// TIA Portal project "交通灯 章家铭" (V15.1)

(* hardware
DEVICE "S7-1200 station_1"  S7-1200 Station
   slot 0: "Rack_0"  S7-1200 Rack  Rack  V1.0
   slot 1: "PLC_1"  CPU 1214C DC/DC/DC  6ES7 214-1AG40-0XB0  V4.2
   slot 2: "DI 16/DQ 16x24VDC_1"  6ES7 223-1BL32-0XB0  V2.0
   slot 3: "AI 4x13BIT/AQ 2x14BIT_1"  6ES7 234-4HE32-0XB0  V2.0
DEVICE "HMI_1"  KTP700 Basic PN
   slot 0: "HMI_1"  KTP700 Basic PN  6AV2 123-2GB03-0AX0  15.1.0.0
   slot 1: "HMI_RT_1"  KTP700 Basic PN  6AV2 123-2GB03-0AX0  15.1.0.0
   slot 5: "HMI_1.IE_CP_1"  PROFINET Interface  15.0.1.0
      slot 1: "PROFINET Interface_1"  PROFINET Interface
         slot 1: "Port_1"  Port
*)

// ===== PLC "PLC_1"  CPU 1214C DC/DC/DC =====

VAR_GLOBAL   // PLC tag table "默认变量表"
   "Tag_1" AT %I8.0 : Bool;
   "Tag_2" AT %I8.1 : Bool;
   "Tag_3" AT %I8.2 : Bool;
   "Tag_4" AT %I8.3 : Bool;
   "Tag_5" AT %I8.4 : Bool;
   "Tag_6" AT %I8.5 : Bool;
   "Tag_7" AT %I8.6 : Bool;
   "Tag_8" AT %I8.7 : Bool;
   "Tag_9" AT %I9.5 : Bool;
   "Tag_10" AT %Q8.0 : Bool;
   "Tag_11" AT %Q8.1 : Bool;
   "Tag_12" AT %Q8.2 : Bool;
   "Tag_13" AT %Q8.3 : Bool;
   "Tag_14" AT %Q8.4 : Bool;
   "Tag_15" AT %Q8.5 : Bool;
   "Tag_16" AT %Q8.6 : Bool;
   "Tag_17" AT %Q8.7 : Bool;
   "Tag_18" AT %Q9.0 : Bool;
   "Tag_19" AT %Q9.1 : Bool;
   "Tag_20" AT %Q9.2 : Bool;
   "Tag_21" AT %Q9.3 : Bool;
   "Tag_22" AT %Q9.4 : Bool;
   "Tag_23" AT %Q9.5 : Bool;
   "Tag_24" AT %Q9.6 : Bool;
   "Tag_25" AT %Q9.7 : Bool;
END_VAR

DATA_BLOCK "code_DB"   // DB1
{ S7_Optimized_Access := 'TRUE' }
VERSION : 0.1
// stored: InstanceOfName code
"code"
BEGIN
END_DATA_BLOCK

FUNCTION_BLOCK "code"   // FB1, SCL
{ S7_Optimized_Access := 'TRUE' }
VERSION : 0.1
   VAR_INPUT
      s01 : Bool;
      s02 : Bool;
      s03 : Bool;
      s04 : Bool;
      s05 : Bool;
      s06 : Bool;
      s07 : Bool;
      s14 : Bool;
   END_VAR
   VAR_OUTPUT
      k01 : Bool;
      k02 : Bool;
      k03 : Bool;
      k04 : Bool;
      k05 : Bool;
      k06 : Bool;
      k07 : Bool;
      k08 : Bool;
      k09 : Bool;
      k10 : Bool;
      k11 : Bool;
      k12 : Bool;
      k13 : Bool;
      k14 : Bool;
      k15 : Bool;
      k16 : Bool;
      hmi_ns_str_time : Int;
      hmi_ns_str_color : Int;
      hmi_ns_left_time : Int;
      hmi_ns_left_color : Int;
      hmi_ew_str_time : Int;
      hmi_ew_str_color : Int;
      hmi_ew_left_color : Int;
      hmi_ew_left_time : Int;
   END_VAR
   VAR
      auto_step : Int;
      ped_active : Bool;
      time_preset : Time;
      timer_auto : TON_TIME;
      timer_ped : TON_TIME;
   END_VAR
   VAR_TEMP
      elapsed_sec : Int;
      t_remain : Int;
      t_ped_remain : Int;
      blink_1hz : Bool;
   END_VAR
BEGIN
   // 初始化
   IF NOT #s01 THEN
       // 钥匙未开启时复位
       #auto_step := 0;
       #ped_active := FALSE;
   ELSE
       // 手动模式
       IF #s02 = TRUE THEN
           // 软件互锁：四个方向的绿灯请求互斥
           #k03 := #s03 AND NOT #s04 AND NOT #s05 AND NOT #s06;
           #k01 := NOT #k03;
           #k02 := FALSE;

           #k06 := #s04 AND NOT #s03 AND NOT #s05 AND NOT #s06;
           #k04 := NOT #k06;
           #k05 := FALSE;

           #k09 := #s05 AND NOT #s03 AND NOT #s04 AND NOT #s06;
           #k07 := NOT #k09;
           #k08 := FALSE;

           #k12 := #s06 AND NOT #s03 AND NOT #s04 AND NOT #s05;
           #k10 := NOT #k12;
           #k11 := FALSE;

           // 自动
       ELSE
           CASE #auto_step OF
               0:
                   #auto_step := 1;

               1:  // 南北直行绿灯
                   #time_preset := T#15s;
                   IF #timer_auto.Q THEN
                       #auto_step := 2;
                   END_IF;

               2:  // 南北直行黄灯
                   #time_preset := T#3s;
                   IF #timer_auto.Q THEN
                       #auto_step := 3;
                   END_IF;

               3:  // 南北左转绿灯
                   #time_preset := T#10s;
                   IF #timer_auto.Q THEN
                       #auto_step := 4;
                   END_IF;

               4:  // 南北左转黄灯
                   #time_preset := T#3s;
                   IF #timer_auto.Q THEN
                       #auto_step := 5;
                   END_IF;

               5:  // 东西直行绿灯
                   #time_preset := T#15s;
                   IF #timer_auto.Q THEN
                       #auto_step := 6;
                   END_IF;

               6:  // 东西直行黄灯
                   #time_preset := T#3s;
                   IF #timer_auto.Q THEN
                       #auto_step := 7;
                   END_IF;

               7:  // 东西左转绿灯
                   #time_preset := T#10s;
                   IF #timer_auto.Q THEN
                       #auto_step := 8;
                   END_IF;

               8:  // 东西左转黄灯
                   #time_preset := T#3s;
                   IF #timer_auto.Q THEN
                       #auto_step := 1;
                   END_IF;

               ELSE
                   #auto_step := 1;
           END_CASE;

           // 驱动自动模式的定时器
           #timer_auto(IN := TRUE,
                       PT := #time_preset);
           IF #timer_auto.Q THEN
               #timer_auto(IN := FALSE,
                           PT := #time_preset);
           END_IF;


           #blink_1hz := ((TIME_TO_DINT(#timer_auto.ET) / 500) MOD 2) = 0;

           #k03 := (#auto_step = 1);
           #k02 := (#auto_step = 2) AND #blink_1hz; 
           #k01 := NOT (#auto_step = 1 OR #auto_step = 2); 

           #k06 := (#auto_step = 3);
           #k05 := (#auto_step = 4) AND #blink_1hz;
           #k04 := NOT (#auto_step = 3 OR #auto_step = 4);

           #k09 := (#auto_step = 5);
           #k08 := (#auto_step = 6) AND #blink_1hz;
           #k07 := NOT (#auto_step = 5 OR #auto_step = 6);

           #k12 := (#auto_step = 7);
           #k11 := (#auto_step = 8) AND #blink_1hz;
           #k10 := NOT (#auto_step = 7 OR #auto_step = 8);


       END_IF;

       // 人行横道控制
       IF #s14 AND NOT #ped_active THEN
           #ped_active := TRUE;
       END_IF;

       // 行人过街定时逻辑
       #timer_ped(IN := #ped_active,
                  PT := T#5s);

       IF #ped_active THEN
           #k14 := FALSE;
           #k13 := TRUE;
           #k16 := FALSE;
           #k15 := TRUE;

           IF #timer_ped.Q THEN
               #ped_active := FALSE;
           END_IF;
       ELSE
           #k14 := TRUE;
           #k13 := FALSE;
           #k16 := TRUE;
           #k15 := FALSE;
       END_IF;

       // ==========================================
       // 5.倒计时
       // 颜色约定: 1=绿灯, 2=黄灯, 3=红灯
       // ==========================================
       IF #s02 THEN
           // 手动模式：没有倒计时(0)，只根据物理绿灯开关状态改变颜色
           #hmi_ns_str_time := 0;
           #hmi_ns_str_color := 3;
           IF #k03 THEN
               #hmi_ns_str_color := 1;
           END_IF;
           #hmi_ns_left_time := 0;
           #hmi_ns_left_color := 3;
           IF #k06 THEN
               #hmi_ns_left_color := 1;
           END_IF;
           #hmi_ew_str_time := 0;
           #hmi_ew_str_color := 3;
           IF #k09 THEN
               #hmi_ew_str_color := 1;
           END_IF;
           #hmi_ew_left_time := 0;
           #hmi_ew_left_color := 3;
           IF #k12 THEN
               #hmi_ew_left_color := 1;
           END_IF;
       ELSE
           // 自动模式：提取当前相位剩余的秒数
           #t_remain := DINT_TO_INT(TIME_TO_DINT(#time_preset) / 1000) - DINT_TO_INT(TIME_TO_DINT(#timer_auto.ET) / 1000);
           IF #t_remain < 0 THEN
               #t_remain := 0;
           END_IF;

           // 核心时间轴投射 (精确计算其他方向等待绿灯的时间)
           CASE #auto_step OF
               1: // 相位: 南北直行绿灯
                   #hmi_ns_str_time := #t_remain;
                   #hmi_ns_str_color := 1; // 绿
                   #hmi_ns_left_time := #t_remain + 3;
                   #hmi_ns_left_color := 3; // 红 (等接下来的黄灯走完)
                   #hmi_ew_str_time := #t_remain + 16;
                   #hmi_ew_str_color := 3; // 红 (3黄+10左+3黄)
                   #hmi_ew_left_time := #t_remain + 34;
                   #hmi_ew_left_color := 3; // 红
               2: // 相位: 南北直行黄灯
                   #hmi_ns_str_time := #t_remain;
                   #hmi_ns_str_color := 2; // 黑
                   #hmi_ns_left_time := #t_remain;
                   #hmi_ns_left_color := 3;
                   #hmi_ew_str_time := #t_remain + 13;
                   #hmi_ew_str_color := 3;
                   #hmi_ew_left_time := #t_remain + 31;
                   #hmi_ew_left_color := 3;
               3: // 相位: 南北左转绿灯
                   #hmi_ns_str_time := #t_remain + 34;
                   #hmi_ns_str_color := 3; // 红
                   #hmi_ns_left_time := #t_remain;
                   #hmi_ns_left_color := 1; // 绿
                   #hmi_ew_str_time := #t_remain + 3;
                   #hmi_ew_str_color := 3;
                   #hmi_ew_left_time := #t_remain + 21;
                   #hmi_ew_left_color := 3;
               4: // 相位: 南北左转黄灯
                   #hmi_ns_str_time := #t_remain + 31;
                   #hmi_ns_str_color := 3;
                   #hmi_ns_left_time := #t_remain;
                   #hmi_ns_left_color := 2; // 黑
                   #hmi_ew_str_time := #t_remain;
                   #hmi_ew_str_color := 3;
                   #hmi_ew_left_time := #t_remain + 18;
                   #hmi_ew_left_color := 3;
               5: // 相位: 东西直行绿灯
                   #hmi_ns_str_time := #t_remain + 16;
                   #hmi_ns_str_color := 3;
                   #hmi_ns_left_time := #t_remain + 34;
                   #hmi_ns_left_color := 3;
                   #hmi_ew_str_time := #t_remain;
                   #hmi_ew_str_color := 1; // 绿
                   #hmi_ew_left_time := #t_remain + 3;
                   #hmi_ew_left_color := 3;
               6: // 相位: 东西直行黄灯
                   #hmi_ns_str_time := #t_remain + 13;
                   #hmi_ns_str_color := 3;
                   #hmi_ns_left_time := #t_remain + 31;
                   #hmi_ns_left_color := 3;
                   #hmi_ew_str_time := #t_remain;
                   #hmi_ew_str_color := 2; // 黑
                   #hmi_ew_left_time := #t_remain;
                   #hmi_ew_left_color := 3;
               7: // 相位: 东西左转绿灯
                   #hmi_ns_str_time := #t_remain + 3;
                   #hmi_ns_str_color := 3;
                   #hmi_ns_left_time := #t_remain + 21;
                   #hmi_ns_left_color := 3;
                   #hmi_ew_str_time := #t_remain + 34;
                   #hmi_ew_str_color := 3;
                   #hmi_ew_left_time := #t_remain;
                   #hmi_ew_left_color := 1; // 绿
               8: // 相位: 东西左转黄灯
                   #hmi_ns_str_time := #t_remain;
                   #hmi_ns_str_color := 3;
                   #hmi_ns_left_time := #t_remain + 18;
                   #hmi_ns_left_color := 3;
                   #hmi_ew_str_time := #t_remain + 31;
                   #hmi_ew_str_color := 3;
                   #hmi_ew_left_time := #t_remain;
                   #hmi_ew_left_color := 2; // 黑
           END_CASE;
       END_IF;



   END_IF;
END_FUNCTION_BLOCK

ORGANIZATION_BLOCK "Main"   // OB1, LAD, ProgramCycle
TITLE = "Main Program Sweep (Cycle)"
{ S7_Optimized_Access := 'TRUE' }
VERSION : 0.1
   VAR_INPUT
      Initial_Call : Bool;   // Initial call of this OB
      Remanence : Bool;   // =True, if remanent data are available
   END_VAR
BEGIN

REGION Network 1
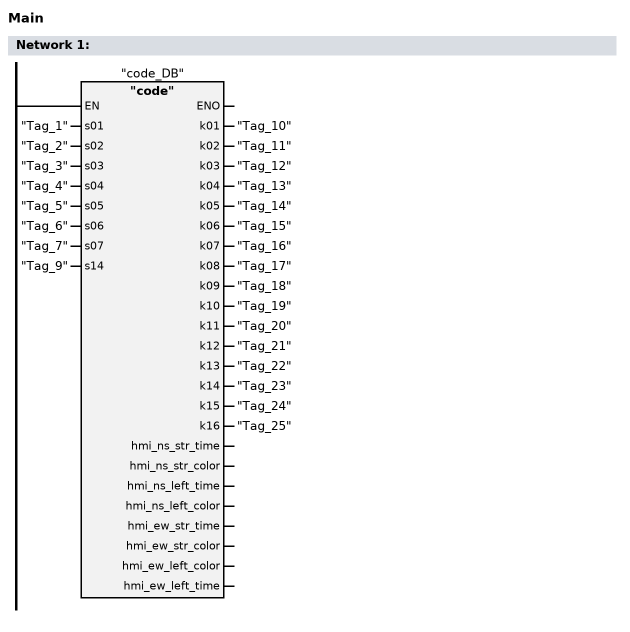
   RUNG wire#powerrail
      "code_DB"(s01 := "Tag_1", s02 := "Tag_2", s03 := "Tag_3", s04 := "Tag_4", s05 := "Tag_5", s06 := "Tag_6", s07 := "Tag_7", s14 := "Tag_9", k01 => "Tag_10", k02 => "Tag_11", k03 => "Tag_12", k04 => "Tag_13", k05 => "Tag_14", k06 => "Tag_15", k07 => "Tag_16", k08 => "Tag_17", k09 => "Tag_18", k10 => "Tag_19", k11 => "Tag_20", k12 => "Tag_21", k13 => "Tag_22", k14 => "Tag_23", k15 => "Tag_24", k16 => "Tag_25", hmi_ns_str_time =>, hmi_ns_str_color =>, hmi_ns_left_time =>, hmi_ns_left_color =>, hmi_ew_str_time =>, hmi_ew_str_color =>, hmi_ew_left_color =>, hmi_ew_left_time =>)
   END_RUNG
   // the same network as SCL:
   "code_DB"(s01 := "Tag_1",   // "code"
             s02 := "Tag_2",
             s03 := "Tag_3",
             s04 := "Tag_4",
             s05 := "Tag_5",
             s06 := "Tag_6",
             s07 := "Tag_7",
             s14 := "Tag_9",
             k01 => "Tag_10",
             k02 => "Tag_11",
             k03 => "Tag_12",
             k04 => "Tag_13",
             k05 => "Tag_14",
             k06 => "Tag_15",
             k07 => "Tag_16",
             k08 => "Tag_17",
             k09 => "Tag_18",
             k10 => "Tag_19",
             k11 => "Tag_20",
             k12 => "Tag_21",
             k13 => "Tag_22",
             k14 => "Tag_23",
             k15 => "Tag_24",
             k16 => "Tag_25");
END_REGION
END_ORGANIZATION_BLOCK

(* ===== HMI "HMI_RT_1" =====
system functions are stored by id; their names below are inferred from use
connection "HMI_连接_1": ETHERNET, SMART_S7_1200_OMS

HMI tags "默认变量表"
   "Tag_ScreenNumber" : UInt, internal
   "code_DB_hmi_ns_str_time" : Int = PLC code_DB.hmi_ns_str_time, 100 ms
   "code_DB_hmi_ns_left_time" : Int = PLC code_DB.hmi_ns_left_time, 100 ms
   "code_DB_hmi_ew_str_time" : Int = PLC code_DB.hmi_ew_str_time, 100 ms
   "code_DB_hmi_ew_left_time" : Int = PLC code_DB.hmi_ew_left_time, 100 ms
   "code_DB_hmi_ns_str_color" : Int = PLC code_DB.hmi_ns_str_color, 100 ms
   "code_DB_hmi_ns_left_color" : Int = PLC code_DB.hmi_ns_left_color, 100 ms
   "code_DB_hmi_ew_str_color" : Int = PLC code_DB.hmi_ew_str_color, 100 ms
   "code_DB_hmi_ew_left_color" : Int = PLC code_DB.hmi_ew_left_color, 100 ms

Template "模板_1" 800x480
   Button "退出" at 714,429 size 71x50; TextOff '退出'; PictureOff "ExitRuntime_KTP700_Basic_PN_TR"; PictureOn "ExitRuntime_KTP700_Basic_PN_TR"
      on Release: StopRuntime(0)
   Button "Template_Button" at 614,429 size 71x50; TextOff 'Text'
   Button "Template_Button_1" at 514,429 size 71x50; TextOff 'Text'
   Button "Template_Button_2" at 414,429 size 71x50; TextOff 'Text'
   Button "Template_Button_3" at 314,429 size 71x50; TextOff 'Text'
   Button "Template_Button_4" at 214,429 size 71x50; TextOff 'Text'
   Button "报警" at 114,429 size 71x50; TextOff '报警'; PictureOff "AlarmDisplay_KTP700_Basic_PN_TR"; PictureOn "AlarmDisplay_KTP700_Basic_PN_TR"
      on Release: function_ef3f5d25("报警窗口_Unacknowledged", -1)
   Button "起始画面" at 14,429 size 71x50; TextOff '起始画面'; PictureOff "NavigateHome_KTP700_Basic_PN_TR"; PictureOn "NavigateHome_KTP700_Basic_PN_TR"
      on Release: ActivateScreen("根画面", 0)
   SymbolicIOField "Symbolic_IO_Field_Screen" at 93,9 size 600x33; TextOff '0'; TextOn '1'; TextList "TextList_ScreenNames"
      ProcessValue <- "Tag_ScreenNumber"
      on Change: ActivateScreenByNumber("Tag_ScreenNumber", 0)
   DateTimeField "HmiScreenItemData" at 695,25 size 105x25
   DateTimeField "HmiScreenItemData_1" at 695,0 size 105x25
   GraphicView "Logo" at 0,0 size 91x51; Picture "HMI_1 的 Logo"

screen "根画面" 800x480, template "模板_1"
   on GenerateScreen: SetTag("Tag_ScreenNumber", 1)
   IOField "I/O 域_1" at 611,160 size 124x94; FormatPattern 99
      ProcessValue <- "code_DB_hmi_ns_str_time"
      Appearance <- "code_DB_hmi_ns_str_color"
   TextField "文本域_1" at 605,122 size 137x37; Text '南北直行'
   IOField "I/O 域_2" at 465,160 size 135x94; FormatPattern 99
      ProcessValue <- "code_DB_hmi_ns_left_time"
      Appearance <- "code_DB_hmi_ns_left_color"
   TextField "文本域_2" at 462,122 size 137x37; Text '南北左转'
   IOField "I/O 域_3" at 200,158 size 123x94; FormatPattern 99
      ProcessValue <- "code_DB_hmi_ew_str_time"
      Appearance <- "code_DB_hmi_ew_str_color"
   TextField "文本域_3" at 192,122 size 137x37; Text '东西直行'
   IOField "I/O 域_4" at 57,158 size 129x94; FormatPattern 99
      ProcessValue <- "code_DB_hmi_ew_left_time"
      Appearance <- "code_DB_hmi_ew_left_color"
   TextField "文本域_4" at 53,122 size 137x37; Text '东西左转'
*)